// TIA Portal V20 export
// export: Created 2026-10-19T18:03:17.5940319Z, ExportSetting WithDefaults, DisplayName Totally Integrated Automation Portal, DisplayVersion V20 Update 6, DisplayName TIA Portal Openness, DisplayVersion V20 Update 6, DisplayName TIA Portal Version Control Interface, DisplayVersion V20 Update 6, DisplayName SINAMICS Startdrive Advanced, DisplayVersion V20 SP1, DisplayName SINAMICS Startdrive G130, G150, S120, S150, SINAMICS MV, G220, S200, S210, DisplayVersion V20 SP1, DisplayName SINAMICS Startdrive G110M, G120, G120C, G120D, G120P, G115D, DisplayVersion V20 SP1, DisplayName STEP 7 Professional, DisplayVersion V20 Update 6, DisplayName STEP 7 Safety, DisplayVersion V20 Update 2, DisplayName WinCC Basic/Comfort/Advanced, DisplayVersion V20 Update 6, DisplayName WinCC Unified, DisplayVersion V20 Update 6
DATA_BLOCK "Order_Table_FB_Carousel_DB"   // DB138
VERSION : 0.1
// stored: AutoNumber true, DBAccessibleFromOPCUA true, DBAccessibleFromWebserver true, InstanceOfName Order_Table_FB_Carousel, InstanceOfType FB
"Order_Table_FB_Carousel"
   // VAR_INPUT
   //    System_Selected { ExternalWritable := 'False'} : Bool;
   //    AutoMan_Switch : Bool;
   //    CurrentTime { ExternalWritable := 'False'} : String;
   //    CurrentDTL : DTL;
   //    Watchdog : "Watchdog_Settings_UDT";
   // END_VAR
   // VAR_IN_OUT
   //    Cnv_Entry : "Inbound_Cnv_Control_UDT";
   //    Cnv_PopUp_1 : "PopUp_Cnv_Control";
   //    WeighingStation : "Stations_DB_UDT";
   //    ProfileStation : "Stations_DB_UDT";
   //    Cnv_PopUp_2 : "PopUp_Cnv_Control";
   //    Cnv_PopUp_3 : "PopUp_Cnv_Control";
   //    Cnv_PopUp_4 : "PopUp_Cnv_Control";
   //    Cnv_Exit : "Outbound_Cnv_Control";
   //    System : "System_UDT";
   //    Control_OPC_Ua : "WMS_OPC_UA";
   // END_VAR
   // VAR
   //    RTR_ITP1_CurrentOrder : UDInt;
   //    RTR_P1P2_CurrentOrder : UDInt;
   //    RTR_P3P4_CurrentOrder : UDInt;
   //    RTR_P4TO_CurrentOrder : UDInt;
   //    Roller_To_Roller_CurrentOrder : UDInt;
   //    Chain_To_Chain_CurrentOrder : UDInt;
   //    Pop4_To_PickSt_CurrentOrder : UDInt;
   //    PickSt_To_Pop1_CurrentOrder : UDInt;
   //    WeighingStation_CurrentOrder { ExternalWritable := 'False'} : UDInt;
   //    ProfileStation_CurrentOrder { ExternalWritable := 'False'} : UDInt;
   //    Roller_To_RollerDoneRTrig : R_TRIG;
   //    RTR_ITP1DoneRTrig { S7_SetPoint := 'True'} : R_TRIG;
   //    RTR_P1P2DoneRTrig { S7_SetPoint := 'True'} : R_TRIG;
   //    RTR_P3P4DoneRTrig { S7_SetPoint := 'True'} : R_TRIG;
   //    RTR_P4TODoneRTrig { S7_SetPoint := 'True'} : R_TRIG;
   //    Chain_To_ChainDoneRTrig : R_TRIG;
   //    Pop4_To_PickSt_DoneRTrig { S7_SetPoint := 'True'} : R_TRIG;
   //    PickSt_To_Pop1_DoneRTrig { S7_SetPoint := 'True'} : R_TRIG;
   //    WeighingStationDoneRTrig { ExternalWritable := 'False'} : R_TRIG;
   //    ProfileStationDoneRTrig { ExternalWritable := 'False'} : R_TRIG;
   //    PalletRefused_1_RTig { ExternalWritable := 'False'} : R_TRIG;
   //    ErrorRTrig { ExternalWritable := 'False'} : R_TRIG;
   //    CancelRTrig { ExternalWritable := 'False'} : R_TRIG;
   //    PauseRTrig { ExternalWritable := 'False'} : R_TRIG;
   //    ResumeRTrig { ExternalWritable := 'False'} : R_TRIG;
   //    Clear_Store : R_TRIG;
   //    Clear_Retrieve : R_TRIG;
   //    Canceling : Bool;
   //    RTR_ITP1_WatchdogTimer : TON_TIME;
   //    RTR_P1P2_WatchdogTimer : TON_TIME;
   //    RTR_P3P4_WatchdogTimer : TON_TIME;
   //    RTR_P4TO_WatchdogTimer : TON_TIME;
   //    Roller_To_Roller_WatchdogTimer { S7_SetPoint := 'True'} : TON_TIME;
   //    Chain_To_Chain_WatchdogTimer { S7_SetPoint := 'True'} : TON_TIME;
   //    Pop4_To_PickWatchdogTimer { S7_SetPoint := 'True'} : TON_TIME;
   //    PickSt_To_Pop1WatchdogTimer : TON_TIME;
   //    WeighingStation_WatchdogTimer : TON_TIME;
   //    ProfileStation_WatchdogTimer : TON_TIME;
   //    Roller_To_Roller_WatchdogStart { S7_SetPoint := 'True'} : Bool;
   //    RTR_ITP1_WatchdogStart : Bool;
   //    RTR_P1P2_WatchdogStart : Bool;
   //    RTR_P3P4_WatchdogStart : Bool;
   //    RTR_P4TO_WatchdogStart : Bool;
   //    Chain_To_Chain_WatchdogStart : Bool;
   //    Pop4_To_PickWatchdogStart : Bool;
   //    PickSt_To_Pop1WatchdogStart : Bool;
   //    WeighingStation_WatchdogStart : Bool;
   //    ProfileStation_WatchdogStart : Bool;
   //    dummy : Int;
   //    dummy_1 : Bool;
   //    dummy_3 : Bool;
   // END_VAR
BEGIN
END_DATA_BLOCK
